(* IEC 61131-3 sources: kns-port-domestic/targets/astra/lib/src/POUs/Base/FB_DeviceBase, 21 files *)

(* ---- FB_DeviceBase.decl.st ---- *)
// Назначение: абстрактная база устройств библиотеки (I_Device, I_AlarmSource): время цикла,
//             режимы (Auto, Manual, Local, OutOfService) с энергонезависимым дистанционным
//             режимом, конфигурация с последней корректной копией (LKG), результат команд,
//             восемь слотов FB_Alarm, сводный статус NAMUR NE 107 и общий заголовок Sts.
//             Тело пустое: порядок цикла задаёт наследник (docs/fb/FB_DeviceBase.md, «Порядок
//             тела»), шаги цикла — защищённые методы. Все переменные секции VAR — часть контракта
//             для наследников, их имена зарезервированы (повтор имени в наследнике — C0097).
// Автор:      kr0nsch
// Версия:     0.1.0
// Документ:   docs/fb/FB_DeviceBase.md
FUNCTION_BLOCK ABSTRACT FB_DeviceBase IMPLEMENTS I_Device
VAR_INPUT
    itfTime : I_TimeSource;                  // источник времени; 0 — встроенный fbSysTime
END_VAR
VAR
    // --- время (BeginCycle) ---
    fbSysTime      : FB_SystemTime;          // запасной источник
    itfTimeAct     : I_TimeSource;           // действующий источник этого вызова
    ltNow          : LTIME;                  // время этого вызова
    ltPrevCall     : LTIME;                  // время предыдущего вызова
    ltDt           : LTIME;                  // ltNow - ltPrevCall; LTIME#0S в первом вызове и при «времени назад»
    xFirstCall     : BOOL := TRUE;           // TRUE до конца первого вызова (FinishCycle)
    // --- режим ---
    eMode          : E_DeviceMode := E_DeviceMode.Manual;   // текущий режим
    xModeReq       : BOOL;                   // есть запрос RequestMode() (снимает FinishCycle)
    eModeReq       : E_DeviceMode := E_DeviceMode.Manual;   // значение запроса; не INT: строгое перечисление (L4)
    stModeMem      : ST_DeviceRetain;        // память режима для ФБ без stRetain (AI, DI)
    xManualIsCheck : BOOL;                   // TRUE у AI/DI: Manual (подмена) даёт CheckFunction
    eDevType       : E_DeviceType := E_DeviceType.None;     // задаёт наследник; FinishCycle пишет в stCommon
    // --- конфигурация ---
    wCfgErr        : WORD;                   // результат CheckConfig этого вызова
    xCfgEverOk     : BOOL;                   // корректная Cfg была хотя бы раз (есть LKG)
    // --- статус ---
    eNe107         : E_Ne107Status := E_Ne107Status.CheckFunction;
    xFault         : BOOL;                   // eNe107 = Failure
    xAvailable     : BOOL;                   // можно рассчитывать на устройство в автомате
    // --- запросы методов ---
    xResetReq      : BOOL;                   // Reset()
    xAckAllReq     : BOOL;                   // AckAll()
    // --- результат команд ---
    eCmdResult     : E_CmdResult := E_CmdResult.None;
    uiCmdSeq       : UINT;                   // +1 на каждую обработанную команду (по кругу)
    // --- тревоги (слоты 0..DEV_ALARMS_MAX - 1) ---
    uiAlarmCount   : UINT;                   // используемых слотов; задаёт наследник в первом вызове
    afbAlarm       : ARRAY[0..GVL_Const.DEV_ALARMS_MAX - 1] OF FB_Alarm;   // слоты тревог
    axAlmCond      : ARRAY[0..GVL_Const.DEV_ALARMS_MAX - 1] OF BOOL;       // условия (заполняет наследник)
    axAlmSuppress  : ARRAY[0..GVL_Const.DEV_ALARMS_MAX - 1] OF BOOL;       // подавление по условию
    arAlmValue     : ARRAY[0..GVL_Const.DEV_ALARMS_MAX - 1] OF REAL;       // значение для события
    wAlmActive     : WORD;                   // бит i: условие слота i активно (после задержек)
    wAlmUnack      : WORD;                   // бит i: слот i не квитирован
    wAlmShelved    : WORD;                   // бит i: слот отложен оператором (Shelved)
    wAlmSuppressed : WORD;                   // бит i: слот подавлен логикой (SuppressedByDesign)
    ePrioUnack     : E_AlarmPriority := E_AlarmPriority.None;   // наивысший приоритет неквитированных
END_VAR

(* ---- AcceptCfg.method.decl.st ---- *)
// Шаг 2 цикла: результат CheckConfig. wErr = 0 — конфигурация корректна: TRUE, вызывающий копирует
// stCfgLkg := stCfg; иначе логика работает по последней корректной копии (LKG)
METHOD PROTECTED AcceptCfg : BOOL
VAR_INPUT
    wErr : WORD;   // биты непройденных проверок (карта wCfgErr устройства)
END_VAR

(* ---- AcceptCfg.method.impl.st ---- *)
wCfgErr := wErr;
IF wErr = 0 THEN
    xCfgEverOk := TRUE;
    AcceptCfg := TRUE;
ELSE
    AcceptCfg := FALSE;
END_IF

(* ---- BeginCycle.method.impl.st ---- *)
ResolveTime();
ltNow := itfTimeAct.Now();
IF NOT xFirstCall AND ltNow >= ltPrevCall THEN
    ltDt := ltNow - ltPrevCall;
ELSE
    // PORT: [types] проверить в Astra.IDE — литералы и преобразования LTIME (C11)
    ltDt := LTIME#0S;
END_IF

(* ---- CheckAlarmCfg.method.decl.st ---- *)
// Проверка конфигурации тревог для CheckConfig устройства: TRUE, если приоритеты всех слотов —
// значения перечисления E_AlarmPriority (0…4)
METHOD PROTECTED CheckAlarmCfg : BOOL
VAR_IN_OUT CONSTANT
    astCfg : ARRAY[0..GVL_Const.DEV_ALARMS_MAX - 1] OF ST_AlarmCfg;   // stCfgIn.astAlarm устройства
END_VAR
VAR
    uiLoop : UINT;                                        // номер слота + 1
    ePrio  : E_AlarmPriority := E_AlarmPriority.Medium;   // приоритет слота
    xOk    : BOOL := TRUE;                                // все проверенные слоты корректны
END_VAR

(* ---- CheckAlarmCfg.method.impl.st ---- *)
FOR uiLoop := 1 TO GVL_Const.DEV_ALARMS_MAX DO
    ePrio := astCfg[uiLoop - 1].ePriority;
    xOk := xOk AND (ePrio = E_AlarmPriority.None OR ePrio = E_AlarmPriority.Low OR ePrio = E_AlarmPriority.Medium
                    OR ePrio = E_AlarmPriority.High OR ePrio = E_AlarmPriority.Critical);
END_FOR
CheckAlarmCfg := xOk;

(* ---- FinishCycle.method.decl.st ---- *)
// Шаг 8 цикла: сводный NE 107 = MAX(статус устройства, статус режима, статус Cfg), Fault, Available,
// общий заголовок stCommon (все 14 полей, старший байт wStatus — общие биты DEV_STS_*), затем
// ltPrevCall := ltNow, конец первого вызова и снятие запросов методов
METHOD PROTECTED FinishCycle
VAR_INPUT
    eDevStatus    : E_Ne107Status;   // статус от логики устройства (Failure, OutOfSpecification, MaintenanceRequired)
    xAvailableDev : BOOL;            // готовность по логике устройства
    wLow          : WORD;            // биты устройства (младший байт wStatus)
    wFaultBits    : WORD;            // wFault
    wWarnBits     : WORD;            // wWarning
END_VAR
VAR_IN_OUT
    stCommon : ST_DeviceSts;         // stSts.stCommon устройства
END_VAR
VAR
    xCfgBad     : BOOL;                                          // нет корректной Cfg или она испорчена
    eModeStatus : E_Ne107Status := E_Ne107Status.Good;           // вклад режима
    eCfgStatus  : E_Ne107Status := E_Ne107Status.Good;           // вклад конфигурации
    wHigh       : WORD;                                          // общие биты 8–15 wStatus
END_VAR

(* ---- FinishCycle.method.impl.st ---- *)
// 1. Сводный статус NE 107 (значения упорядочены по тяжести: MAX). Режим даёт CheckFunction: OutOfService, подмена
//    AI/DI (Manual) и Local — механизмом управляют по месту, выход ПЛК не действует (категория C NE 107, статус PA
//    «function check / local override», NE107-1)
xCfgBad := wCfgErr <> 0 OR NOT xCfgEverOk;
IF eMode = E_DeviceMode.OutOfService OR eMode = E_DeviceMode.Local
   OR (xManualIsCheck AND eMode = E_DeviceMode.Manual)
THEN
    eModeStatus := E_Ne107Status.CheckFunction;
END_IF
IF xCfgBad THEN
    eCfgStatus := E_Ne107Status.CheckFunction;
END_IF
eNe107 := F_Ne107Worst(eA := eDevStatus, eB := eModeStatus);
eNe107 := F_Ne107Worst(eA := eNe107, eB := eCfgStatus);
xFault := eNe107 = E_Ne107Status.Failure;
xAvailable := xAvailableDev AND xCfgEverOk;

// 2. Общий старший байт wStatus (раздел 5.2 контракта)
IF eMode = E_DeviceMode.Auto THEN
    wHigh := wHigh OR GVL_Const.DEV_STS_MODE_AUTO;
ELSIF eMode = E_DeviceMode.Manual THEN
    wHigh := wHigh OR GVL_Const.DEV_STS_MODE_MANUAL;
ELSIF eMode = E_DeviceMode.Local THEN
    wHigh := wHigh OR GVL_Const.DEV_STS_MODE_LOCAL;
ELSIF eMode = E_DeviceMode.OutOfService THEN
    wHigh := wHigh OR GVL_Const.DEV_STS_MODE_OOS;
END_IF
IF xCfgBad THEN
    wHigh := wHigh OR GVL_Const.DEV_STS_CFG_ERROR;
END_IF
IF xFault THEN
    wHigh := wHigh OR GVL_Const.DEV_STS_FAILURE;
END_IF
IF wWarnBits <> 0 OR eNe107 = E_Ne107Status.OutOfSpecification
   OR eNe107 = E_Ne107Status.MaintenanceRequired
THEN
    wHigh := wHigh OR GVL_Const.DEV_STS_WARNING;
END_IF
IF wAlmUnack <> 0 THEN
    wHigh := wHigh OR GVL_Const.DEV_STS_ALARM_UNACK;
END_IF

// 3. Общий заголовок состояния
stCommon.wStatus := (wLow AND GVL_Const.WORD_LOW_BYTE) OR wHigh;
stCommon.wFault := wFaultBits;
stCommon.wWarning := wWarnBits;
stCommon.wCfgErr := wCfgErr;
stCommon.eMode := eMode;
stCommon.eNe107 := eNe107;
stCommon.eCmdResult := eCmdResult;
stCommon.uiCmdSeq := uiCmdSeq;
stCommon.wAlmActive := wAlmActive;
stCommon.wAlmUnack := wAlmUnack;
stCommon.wAlmShelved := wAlmShelved;
stCommon.ePrioUnack := ePrioUnack;
stCommon.eDevType := eDevType;
stCommon.wAlmSuppressed := wAlmSuppressed;

// 4. Конец цикла
ltPrevCall := ltNow;
xFirstCall := FALSE;
xResetReq := FALSE;
xAckAllReq := FALSE;
xModeReq := FALSE;

(* ---- GetAlarm.method.decl.st ---- *)
// Тревога слота uiIndex через интерфейс; вне 0..AlarmCount - 1 — 0
METHOD PUBLIC GetAlarm : I_Alarm
VAR_INPUT
    uiIndex : UINT;   // номер слота
END_VAR

(* ---- GetAlarm.method.impl.st ---- *)
IF uiIndex < MIN(uiAlarmCount, GVL_Const.DEV_ALARMS_MAX) THEN
    GetAlarm := afbAlarm[uiIndex];
ELSE
    GetAlarm := 0;
END_IF

(* ---- OnModeChanged.method.decl.st ---- *)
// Виртуальный хук смены режима, в базе пуст. Вызывается только как THIS^.OnModeChanged(...) из
// ProcessMode и SwitchRemoteMode, в том числе в первом вызове, если режим из stRetain отличается
// от начального Manual (наследник отличает этот случай по xFirstCall). Наследник переопределяет с
// той же сигнатурой и PROTECTED и в начале вызывает SUPER^.OnModeChanged(eOld := eOld, eNew := eNew).
// Хук НЕ ДОЛЖЕН трогать VAR_IN_OUT устройства (R2)
METHOD PROTECTED OnModeChanged
VAR_INPUT
    eOld : E_DeviceMode;   // режим до смены
    eNew : E_DeviceMode;   // новый режим
END_VAR

(* ---- ProcessMode.method.decl.st ---- *)
// Шаг 4 цикла: автомат режима. Санитизация stRetain.eRemoteMode; победивший запрос среди битов
// stCmd и RequestMode() по старшинству OutOfService > Manual > Auto (одновременные запросы —
// одна команда); сброс импульсов режима; новый режим по старшинству OutOfService > Local >
// дистанционный; при смене — виртуальный хук THIS^.OnModeChanged. Результат None — запросов не было
METHOD PROTECTED ProcessMode : E_CmdResult
VAR_INPUT
    xLocalSel       : BOOL;   // переключатель в положении «Местное»
    xLocalSupported : BOOL;   // у типа есть режим Local
    xOosAllowed     : BOOL;   // механизм стоит: вывод из работы допустим
END_VAR
VAR_IN_OUT
    stCmd    : ST_DeviceCmd;      // общий заголовок команд: импульсы режима сбрасываются
    stRetain : ST_DeviceRetain;   // дистанционный режим и признак OutOfService (AI/DI — stModeMem)
END_VAR
VAR
    xAnyReq   : BOOL;                                    // в этом вызове есть запрос режима
    eWinner   : E_DeviceMode := E_DeviceMode.Manual;     // победивший запрос
    eModeOld  : E_DeviceMode := E_DeviceMode.Manual;     // режим до смены
    eModeNew  : E_DeviceMode := E_DeviceMode.Manual;     // режим по итогам вызова
    eResult   : E_CmdResult := E_CmdResult.None;         // результат запроса режима
END_VAR

(* ---- ProcessMode.method.impl.st ---- *)
// 1. Санитизация: значение вне {Auto, Manual} (0 после очистки, мусор persistent-памяти) — Manual.
//    Строгое перечисление защищает только исходный текст, поэтому проверка — сравнениями
IF stRetain.eRemoteMode <> E_DeviceMode.Auto AND stRetain.eRemoteMode <> E_DeviceMode.Manual THEN
    stRetain.eRemoteMode := E_DeviceMode.Manual;
END_IF

// 2. Победивший запрос: биты stCmd и RequestMode() вместе, по старшинству OutOfService > Manual > Auto
xAnyReq := TRUE;
IF stCmd.xSetOos OR (xModeReq AND eModeReq = E_DeviceMode.OutOfService) THEN
    eWinner := E_DeviceMode.OutOfService;
ELSIF stCmd.xSetManual OR (xModeReq AND eModeReq = E_DeviceMode.Manual) THEN
    eWinner := E_DeviceMode.Manual;
ELSIF stCmd.xSetAuto OR (xModeReq AND eModeReq = E_DeviceMode.Auto) THEN
    eWinner := E_DeviceMode.Auto;
ELSE
    xAnyReq := FALSE;
END_IF
stCmd.xSetAuto := FALSE;
stCmd.xSetManual := FALSE;
stCmd.xSetOos := FALSE;
xModeReq := FALSE;

// 3. Выполнение: OutOfService — только при стоящем механизме (повтор в OutOfService принимается);
//    Auto и Manual запоминаются в stRetain (в Local тоже) и выводят из OutOfService
IF xAnyReq THEN
    IF eWinner = E_DeviceMode.OutOfService THEN
        IF xOosAllowed OR stRetain.xOutOfService THEN
            stRetain.xOutOfService := TRUE;
            eResult := E_CmdResult.Accepted;
        ELSE
            eResult := E_CmdResult.RejectedState;
        END_IF
    ELSE
        stRetain.eRemoteMode := eWinner;
        stRetain.xOutOfService := FALSE;
        eResult := E_CmdResult.Accepted;
    END_IF
END_IF
ProcessMode := eResult;

// 4. Режим по старшинству OutOfService > Local > дистанционный
IF stRetain.xOutOfService THEN
    eModeNew := E_DeviceMode.OutOfService;
ELSIF xLocalSel AND xLocalSupported THEN
    eModeNew := E_DeviceMode.Local;
ELSE
    eModeNew := stRetain.eRemoteMode;
END_IF
IF eModeNew <> eMode THEN
    eModeOld := eMode;
    eMode := eModeNew;
    THIS^.OnModeChanged(eOld := eModeOld, eNew := eModeNew);
END_IF

(* ---- RequestMode.method.decl.st ---- *)
// Запрос режима для станционной логики, как бит stCmd: Auto, Manual, OutOfService — TRUE (запрос
// выполнит ProcessMode ближайшего вызова, результат — в eCmdResult); Local и прочее — FALSE.
// Имя параметра не eMode: оно затенило бы переменную базы (L3)
METHOD PUBLIC RequestMode : BOOL
VAR_INPUT
    eNewMode : E_DeviceMode;   // требуемый режим
END_VAR

(* ---- RequestMode.method.impl.st ---- *)
IF eNewMode = E_DeviceMode.Auto OR eNewMode = E_DeviceMode.Manual OR eNewMode = E_DeviceMode.OutOfService THEN
    eModeReq := eNewMode;
    xModeReq := TRUE;
    RequestMode := TRUE;
ELSE
    RequestMode := FALSE;
END_IF

(* ---- ResolveTime.method.impl.st ---- *)
IF itfTime <> 0 THEN
    itfTimeAct := itfTime;
ELSE
    itfTimeAct := fbSysTime;
END_IF

(* ---- RunAlarms.method.decl.st ---- *)
// Шаг 7 цикла: запросы тревог (квитировать всё, маски квитирования, shelve и unshelve), вызов
// используемых слотов и сводка wAlmActive, wAlmUnack, wAlmShelved, wAlmSuppressed, ePrioUnack. Сбрасывает xAck,
// xReset и маски stCmd. Циклы — FOR uiLoop := 1 TO MIN(uiAlarmCount, DEV_ALARMS_MAX): при 0 слотов
// беззнаковое «uiAlarmCount - 1» не возникает
METHOD PROTECTED RunAlarms
VAR_INPUT
    udiIdBase : UDINT;            // номер первой тревоги устройства (stCfgLkg.udiAlarmIdBase)
END_VAR
VAR_IN_OUT
    stCmd : ST_DeviceCmd;         // общий заголовок команд
END_VAR
VAR_IN_OUT CONSTANT
    astCfg : ARRAY[0..GVL_Const.DEV_ALARMS_MAX - 1] OF ST_AlarmCfg;   // stCfgLkg.astAlarm
END_VAR
VAR
    uiUsed     : UINT;            // слотов в работе: MIN(uiAlarmCount, DEV_ALARMS_MAX)
    uiLoop     : UINT;            // номер слота + 1
    uiSlot     : UINT;            // номер слота
    wBit       : WORD;            // бит слота в масках
    xAckAllNow : BOOL;            // квитировать все слоты
    xShelveAny : BOOL;            // хотя бы один слот принял shelve
    xAccepted  : BOOL;            // ответ метода слота (запрос выполнит вызов слота ниже)
    eSlotState : E_AlarmState := E_AlarmState.Normal;   // состояние слота
END_VAR

(* ---- RunAlarms.method.impl.st ---- *)
uiUsed := MIN(uiAlarmCount, GVL_Const.DEV_ALARMS_MAX);

// 1. Запросы: квитировать всё (xAck, xReset, AckAll(), Reset()), маски по слотам. Методы слотов
//    только ставят запрос — его выполняет вызов слота в шаге 2 этого же цикла
xAckAllNow := stCmd.xAck OR stCmd.xReset OR xAckAllReq OR xResetReq;
FOR uiLoop := 1 TO uiUsed DO
    uiSlot := uiLoop - 1;
    wBit := SHL(WORD#16#0001, uiSlot);
    IF xAckAllNow OR (stCmd.wAckReq AND wBit) <> 0 THEN
        xAccepted := afbAlarm[uiSlot].Ack();
    END_IF
    // в OutOfService shelve не принимается (10.1); проверка по режиму устройства, а не по ответу
    // слота: в вызове входа в OutOfService слот ещё не в OutOfService и ответил бы TRUE, а его тело
    // запрос отклонит — результат команды был бы ложным Accepted
    IF (stCmd.wShelveReq AND wBit) <> 0 AND eMode <> E_DeviceMode.OutOfService THEN
        xAccepted := afbAlarm[uiSlot].Shelve(tDuration := T#0S);
        xShelveAny := xShelveAny OR xAccepted;
    END_IF
    IF (stCmd.wUnshelveReq AND wBit) <> 0 THEN
        xAccepted := afbAlarm[uiSlot].Unshelve();
    END_IF
END_FOR
// результаты: «квитировать всё» (xAck и AckAll() вместе — одна команда) и каждая ненулевая маска;
// xReset и Reset() дают результат в шаге Reset устройства
IF stCmd.xAck OR xAckAllReq THEN
    SetCmdResult(eResult := E_CmdResult.Accepted);
END_IF
IF stCmd.wAckReq <> 0 THEN
    SetCmdResult(eResult := E_CmdResult.Accepted);
END_IF
IF stCmd.wShelveReq <> 0 THEN
    IF xShelveAny THEN
        SetCmdResult(eResult := E_CmdResult.Accepted);
    ELSE
        SetCmdResult(eResult := E_CmdResult.RejectedState);
    END_IF
END_IF
IF stCmd.wUnshelveReq <> 0 THEN
    SetCmdResult(eResult := E_CmdResult.Accepted);
END_IF
stCmd.xAck := FALSE;
stCmd.xReset := FALSE;
stCmd.wAckReq := 0;
stCmd.wShelveReq := 0;
stCmd.wUnshelveReq := 0;

// 2. Вызов слотов и 3. сводка. OutOfService устройства — OutOfService у всех слотов
wAlmActive := 0;
wAlmUnack := 0;
wAlmShelved := 0;
wAlmSuppressed := 0;
ePrioUnack := E_AlarmPriority.None;
FOR uiLoop := 1 TO uiUsed DO
    uiSlot := uiLoop - 1;
    wBit := SHL(WORD#16#0001, uiSlot);
    afbAlarm[uiSlot](xIn := axAlmCond[uiSlot], xSuppress := axAlmSuppress[uiSlot],
                     xOutOfService := (eMode = E_DeviceMode.OutOfService), udiId := udiIdBase + uiSlot,
                     rValue := arAlmValue[uiSlot], stCfg := astCfg[uiSlot], itfTime := itfTimeAct);
    IF afbAlarm[uiSlot].Active THEN
        wAlmActive := wAlmActive OR wBit;
    END_IF
    IF afbAlarm[uiSlot].Unacked THEN
        wAlmUnack := wAlmUnack OR wBit;
        ePrioUnack := MAX(ePrioUnack, afbAlarm[uiSlot].AlarmPriority);
    END_IF
    // наложенные состояния ISA-18.2 — раздельно (ALM-2): отложенные оператором (список отложенных тревог с
    // остатком срока) и подавленные логикой; OutOfService слотов совпадает с режимом устройства (eMode)
    eSlotState := afbAlarm[uiSlot].State;
    IF eSlotState = E_AlarmState.Shelved THEN
        wAlmShelved := wAlmShelved OR wBit;
    ELSIF eSlotState = E_AlarmState.SuppressedByDesign THEN
        wAlmSuppressed := wAlmSuppressed OR wBit;
    END_IF
END_FOR

(* ---- SetCmdResult.method.decl.st ---- *)
// Результат обработанной команды: eCmdResult и uiCmdSeq + 1 (UINT, по кругу)
METHOD PROTECTED SetCmdResult
VAR_INPUT
    eResult : E_CmdResult;   // результат команды
END_VAR

(* ---- SwitchRemoteMode.method.decl.st ---- *)
// Смена дистанционного режима логикой устройства («Стоп» в Auto → Manual, снятие подмены AI/DI по
// времени, ПИД ShedToManual): запоминается в stRetain; если устройство в дистанционном режиме —
// режим меняется сразу, с хуком THIS^.OnModeChanged. Значения кроме Auto и Manual не принимаются
METHOD PROTECTED SwitchRemoteMode
VAR_INPUT
    eNew : E_DeviceMode;          // Auto или Manual
END_VAR
VAR_IN_OUT
    stRetain : ST_DeviceRetain;   // дистанционный режим (AI/DI — stModeMem)
END_VAR
VAR
    eModeOld : E_DeviceMode := E_DeviceMode.Manual;   // режим до смены
END_VAR

(* ---- SwitchRemoteMode.method.impl.st ---- *)
IF eNew = E_DeviceMode.Auto OR eNew = E_DeviceMode.Manual THEN
    stRetain.eRemoteMode := eNew;
    IF (eMode = E_DeviceMode.Auto OR eMode = E_DeviceMode.Manual) AND eMode <> eNew THEN
        eModeOld := eMode;
        eMode := eNew;
        THIS^.OnModeChanged(eOld := eModeOld, eNew := eNew);
    END_IF
END_IF
